DATA_BLOCK "naut_SfcStepMaxtime_DB"
{ S7_Optimized_Access := 'TRUE' }
VERSION : 0.1
"naut_SfcStepMaxtime"

BEGIN

END_DATA_BLOCK
